(* IEC 61131-3 sources: conveyor-codesys-oop/src, 4 files *)

(* ---- E_State.st ---- *)
TYPE E_State :
(
    IDLE       := 0,   // Waiting for start command
    RUNNING    := 1,   // Conveyor running, counting products
    BATCH_DONE := 2,   // Target count reached, waiting for reset
    ESTOP      := 3    // Emergency stop active, latched until reset
);
END_TYPE

(* ---- FB_Conveyor.st ---- *)
// --- Declaration ---
FUNCTION_BLOCK FB_Conveyor IMPLEMENTS IConveyor
VAR_INPUT
    bSensor   : BOOL;           // Product detection sensor
    bEStopNC  : BOOL := TRUE;   // Emergency stop (NC: TRUE in normal condition)
    iTarget   : INT := 10;      // Target count per batch
END_VAR
VAR_OUTPUT
    bMotor       : BOOL;        // Conveyor motor
    bBatchDone   : BOOL;        // TRUE when the batch is complete
    bEStopActive : BOOL;        // TRUE while in emergency stop state
    iCount       : INT;         // Product counter
END_VAR
VAR
    eState    : E_State := E_State.IDLE;   // Current machine state
    rtSensor  : R_TRIG;                    // Rising edge detector for the sensor

    // Command requests, set by the methods and cleared at the end of each cycle
    bStartReq : BOOL;
    bStopReq  : BOOL;
    bResetReq : BOOL;
END_VAR

// --- Implementation ---
// Detect rising edge of the sensor (one pulse per product)
rtSensor(CLK := bSensor);

// E-Stop has priority over everything, in every state
IF NOT bEStopNC THEN
    eState := E_State.ESTOP;
END_IF

CASE eState OF

    E_State.IDLE:
        bMotor := FALSE;
        // Start is ignored if a stop request arrives in the same cycle
        IF bStartReq AND NOT bStopReq THEN
            iCount := 0;
            eState := E_State.RUNNING;
        END_IF

    E_State.RUNNING:
        bMotor := TRUE;
        IF rtSensor.Q THEN
            iCount := iCount + 1;
        END_IF
        IF bStopReq THEN
            // Normal stop: back to idle
            eState := E_State.IDLE;
        ELSIF iCount >= iTarget THEN
            // Batch finished
            eState := E_State.BATCH_DONE;
        END_IF

    E_State.BATCH_DONE:
        bMotor := FALSE;
        IF bResetReq THEN
            iCount := 0;
            eState := E_State.IDLE;
        END_IF

    E_State.ESTOP:
        bMotor := FALSE;
        // E-Stop must be released AND a reset request is required
        IF bEStopNC AND bResetReq THEN
            iCount := 0;
            eState := E_State.IDLE;
        END_IF

END_CASE

// Status outputs are driven directly from the current state
bBatchDone   := (eState = E_State.BATCH_DONE);
bEStopActive := (eState = E_State.ESTOP);

// Clear the requests: each method call is valid for one cycle only
bStartReq := FALSE;
bStopReq  := FALSE;
bResetReq := FALSE;

// ===== Method: Start =====
METHOD Start
// Request a start (valid for one cycle)
bStartReq := TRUE;

// ===== Method: Stop =====
METHOD Stop
// Request a normal stop (valid for one cycle)
bStopReq := TRUE;

// ===== Method: Reset =====
METHOD Reset
// Request a reset after batch complete or emergency stop (valid for one cycle)
bResetReq := TRUE;

(* ---- FB_JamConveyor.st ---- *)
// --- Declaration ---
FUNCTION_BLOCK FB_JamConveyor EXTENDS FB_Conveyor
VAR_INPUT
    tJamTimeout : TIME := T#5S;   // Max time without a product while running
END_VAR
VAR_OUTPUT
    bJam : BOOL;                  // TRUE when a jam has been detected
END_VAR
VAR
    tonJam : TON;                 // Timer for jam detection
END_VAR

// --- Implementation ---
// Run the base class logic first (not called automatically in CODESYS)
SUPER^();

// Jam detection: motor running but no product detected for tJamTimeout.
// The timer is reset by every product (rising edge of the sensor).
tonJam(IN := (eState = E_State.RUNNING) AND NOT rtSensor.Q, PT := tJamTimeout);

IF tonJam.Q THEN
    bJam := TRUE;
    eState := E_State.IDLE;   // Stop the conveyor
END_IF

// Status outputs are driven directly from the current state
bBatchDone   := (eState = E_State.BATCH_DONE);
bEStopActive := (eState = E_State.ESTOP);

// Clear the requests: each method call is valid for one cycle only
bStartReq := FALSE;
bStopReq  := FALSE;
bResetReq := FALSE;

// ===== Method: Start =====
METHOD Start
// Override: ignore start requests while a jam is active
IF NOT bJam THEN
    SUPER^.Start();   // Call the base class method
END_IF

// ===== Method: Reset =====
METHOD Reset
// Override: also clear the jam flag, then do the normal reset
bJam := FALSE;
SUPER^.Reset();

(* ---- PLC_PRG.st ---- *)
PROGRAM PLC_PRG
VAR
    // --- Inputs (bound to the visualization) ---
    bStart    : BOOL;           // Start button (NO)
    bStopNC   : BOOL := TRUE;   // Stop button (NC)
    bEStopNC  : BOOL := TRUE;   // Emergency stop (NC)
    bReset    : BOOL;           // Reset button (NO)
    bSensor   : BOOL;           // Sensor of conveyor 1
    bSensor2  : BOOL;           // Sensor of conveyor 2 (test via watch window)

    // --- Outputs of conveyor 1 (bound to the visualization) ---
    bMotor     : BOOL;
    bBatchLamp : BOOL;
    bEStopLamp : BOOL;
    iCount     : INT;

    // --- Edge detectors for the buttons ---
    rtStart   : R_TRIG;
    rtReset   : R_TRIG;

    // --- Two instances: one base type, one derived type ---
    Conv1     : FB_Conveyor;
    Conv2     : FB_JamConveyor := (iTarget := 5);   // different batch size

    // --- Interface references for polymorphic access ---
    aConv     : ARRAY[1..2] OF IConveyor;
    i         : INT;

    // --- Mirror of conveyor 2 outputs, for easy monitoring ---
    bMotor2   : BOOL;
    bJam2     : BOOL;
END_VAR

// Edge detection for the buttons
rtStart(CLK := bStart);
rtReset(CLK := bReset);

// Bind interface references to the concrete instances
aConv[1] := Conv1;
aConv[2] := Conv2;

// Polymorphic commands: the loop does not know which type each element is
FOR i := 1 TO 2 DO
    IF rtStart.Q THEN
        aConv[i].Start();
    END_IF
    IF NOT bStopNC THEN
        aConv[i].Stop();
    END_IF
    IF rtReset.Q THEN
        aConv[i].Reset();
    END_IF
END_FOR

// Cyclic execution of each instance
Conv1(bSensor := bSensor,  bEStopNC := bEStopNC);
Conv2(bSensor := bSensor2, bEStopNC := bEStopNC, tJamTimeout := T#5S);

// Map conveyor 1 outputs to the variables used by the visualization
bMotor     := Conv1.bMotor;
bBatchLamp := Conv1.bBatchDone;
bEStopLamp := Conv1.bEStopActive;
iCount     := Conv1.iCount;

// Mirror conveyor 2 outputs
bMotor2 := Conv2.bMotor;
bJam2   := Conv2.bJam;
